FUNCTION_BLOCK FB_LightTower
VAR_INPUT
	bBuzzerBypass: BOOL;
END_VAR
VAR_OUTPUT
	qLedGreen	: BOOL;
	qLedYellow	: BOOL;
	qLedRed		: BOOL;
	qLedBlue	: BOOL;
	qBuzzer		: BOOL;		
	
	qSignal_1: BOOL; //wire BN
	qSignal_2: BOOL; //wire GY
	qSignal_3: BOOL; //wire BK
	qSignal_4: BOOL; //wire WT

END_VAR
VAR
	eLightTowerState		: E_LightTowerState;
	eLightTower_Type		: E_LightTower_Type:=E_LightTower_Type.eSingleLayer;

	
	ton_Blink				: TON;
	ton_Buzzer				: TON;
	t_Buzzer				: TIME:=T#2S;
	t_BuzzerShort			: TIME:=T#0.5S;
	t_BuzzerErrorDelay		: TIME:=T#10S;
	t_BuzzerWarningDelay	: TIME:=T#30S;
	//eLightTowerState_Last	: E_LightTowerState;
	bBuzzerMuteMemo: BOOL;	
	ton_MuteBuzzer: TON;
	ton_NoMessage: TON;
	ton_BuzzerLongTimeOn: TON;	
END_VAR

ton_Blink(IN:=NOT ton_Blink.Q);
CASE eLightTower_Type OF
	E_LightTower_Type.eSingleLayer: m_Single_Layer();
	E_LightTower_Type.eMultiLayer: m_Multi_Layer();
	
END_CASE


ton_NoMessage(PT:=T#5S,IN:=bBuzzerMuteMemo AND iActErrors=0 AND iActWarning=0);

IF (stOpMain.bSetPlay
	(*OR stOpLoad.bSetPlay
	OR stOpUnload.bSetPlay
	OR stOpManip.bSetPlay
	OR stOpHMI.bSetPlay
	OR prg_Call_OpMode.fbModeIndex.rt_Play.Q
	OR prg_Call_OpMode.fbModeLoad.rt_Play.Q
	OR prg_Call_OpMode.fbModeUnload.rt_Play.Q
	OR prg_Call_OpMode.fbModeManip.rt_Play.Q*)
	OR ton_NoMessage.Q	
)
THEN;
	ton_MuteBuzzer.IN:=TRUE;
END_IF
IF ton_MuteBuzzer.IN THEN;
	bBuzzerMuteMemo:=FALSE;
END_IF
ton_MuteBuzzer(PT:=T#1S);
IF ton_MuteBuzzer.Q THEN
	ton_MuteBuzzer.IN:=FALSE;
END_IF
IF prg_Messages.ResetErrors OR ton_BuzzerLongTimeOn.Q THEN;// iActErrors=0 AND iActWarning=0
	bBuzzerMuteMemo:=TRUE;
END_IF
ton_BuzzerLongTimeOn(PT:=T#30M,IN:=eBuzzerMode<>eBuzzerOff);

(*
TYPE E_BuzzerMode :
(
	eBuzzerOff := 0,
	eBuzzerError,		//Short Delay Off
	eBuzzerWarning		//Long Delay Off
);
END_TYPE
*)

IF NOT bBuzzerBypass THEN
	ton_Buzzer();
	CASE eBuzzerMode OF
		eBuzzerOff :;
			qBuzzer:=FALSE;
			
			ton_Buzzer.IN:=FALSE;
		eBuzzerError:;			//Short Delay Off
			qBuzzer:=TRUE;
			ton_Buzzer.PT:=t_BuzzerErrorDelay;
			ton_Buzzer.IN:=NOT ton_Buzzer.Q;
			IF ton_Buzzer.ET>t_Buzzer THEN; qBuzzer:=FALSE; END_IF
		eBuzzerWarning:;		//Long Delay Off
			qBuzzer:=TRUE;
			ton_Buzzer.PT:=t_BuzzerWarningDelay;
			ton_Buzzer.IN:=NOT ton_Buzzer.Q;
			IF ton_Buzzer.ET>t_BuzzerShort THEN; qBuzzer:=FALSE; END_IF
	END_CASE	
ELSE
	qBuzzer:=FALSE;
END_IF

METHOD m_Multi_Layer : BOOL
VAR_INPUT
END_VAR
CASE eLightTowerState OF
	E_LightTowerState.eLightsOff:;
		qLedGreen	:=FALSE;
		qLedYellow	:=FALSE;
		qLedRed		:=FALSE;
		qLedBlue	:=FALSE;
		eBuzzerMode:=eBuzzerOff;	
		
	E_LightTowerState.eGreen:;
		qLedGreen	:=TRUE;
		qLedYellow	:=FALSE;
		qLedRed		:=FALSE;
		qLedBlue	:=FALSE;
		eBuzzerMode:=eBuzzerOff;	
		
	E_LightTowerState.eGreen_YellowBlink:;
		qLedGreen	:=TRUE;
		qLedYellow	:=TRUE;
		qLedRed		:=FALSE;
		qLedBlue	:=FALSE;
		IF bBuzzerMuteMemo THEN;
			eBuzzerMode:=eBuzzerOff;
		ELSE
			eBuzzerMode:=eBuzzerWarning;
		END_IF
		ton_Blink.PT:=T#1S;
		IF ton_Blink.ET>T#0.5S THEN; qLedYellow:=FALSE; ELSE;qLedGreen:=FALSE; END_IF	
		
	E_LightTowerState.eGreenBlink:;
		qLedGreen	:=TRUE;
		qLedYellow	:=FALSE;
		qLedRed		:=FALSE;
		qLedBlue	:=FALSE;
		eBuzzerMode:=eBuzzerOff;		
		ton_Blink.PT:=T#1S;
		IF ton_Blink.ET>T#0.5S THEN; qLedGreen:=FALSE; END_IF	

	E_LightTowerState.eGreenBlink_YellowBlink:;
		qLedGreen	:=TRUE;
		qLedYellow	:=TRUE;
		qLedRed		:=FALSE;
		qLedBlue	:=FALSE;
		IF bBuzzerMuteMemo THEN;
			eBuzzerMode:=eBuzzerOff;
		ELSE
			eBuzzerMode:=eBuzzerWarning;
		END_IF
		ton_Blink.PT:=T#1S;
		IF ton_Blink.ET>T#0.5S THEN; qLedYellow:=FALSE; ELSE;qLedGreen:=FALSE; END_IF

	E_LightTowerState.eGreenBlink_RedBlink:;
		qLedGreen	:=TRUE;
		qLedYellow	:=FALSE;
		qLedRed		:=TRUE;
		qLedBlue	:=FALSE;
		IF bBuzzerMuteMemo THEN;
			eBuzzerMode:=eBuzzerOff;
		ELSE
			eBuzzerMode:=eBuzzerError;
		END_IF
		ton_Blink.PT:=T#1S;
		IF ton_Blink.ET>T#0.5S THEN; qLedRed:=FALSE; ELSE;qLedGreen:=FALSE; END_IF
		
	E_LightTowerState.eYellow:;
		qLedGreen	:=FALSE;
		qLedYellow	:=TRUE;
		qLedRed		:=FALSE;
		qLedBlue	:=FALSE;
		eBuzzerMode:=eBuzzerOff;	
		
	E_LightTowerState.eRed:;
		qLedGreen	:=FALSE;
		qLedYellow	:=FALSE;
		qLedRed		:=TRUE;
		qLedBlue	:=FALSE;
		IF bBuzzerMuteMemo THEN;
			eBuzzerMode:=eBuzzerOff;
		ELSE
			eBuzzerMode:=eBuzzerError;
		END_IF
		
	E_LightTowerState.eBlue:;
		qLedGreen	:=FALSE;
		qLedYellow	:=FALSE;
		qLedRed		:=FALSE;
		qLedBlue	:=TRUE;
		eBuzzerMode:=eBuzzerOff;	
				
END_CASE
END_METHOD

METHOD m_Op_Case1 : BOOL
VAR_INPUT
END_VAR
IF 		stOpMain.iActOperation=E_OperationButtons.ePauseAll
	AND iActErrors<>0
	THEN;	
	eLightTowerState:=E_LightTowerState.eRed;
 						//7
ELSIF 	stOpMain.iActOperation=E_OperationButtons.ePauseAll
	AND iActErrors=0
	THEN;
	eLightTowerState:=E_LightTowerState.eYellow;					//6	
	
ELSIF 	stOpMain.iActOperation=E_OperationButtons.ePlayAll
	AND iActErrors=0
 	AND iActWarning<>0
	THEN;
	eLightTowerState:=E_LightTowerState.eGreenBlink_YellowBlink;	//4
		
ELSIF 	stOpMain.iActOperation=E_OperationButtons.ePlayAll
	AND iActErrors=0 
	AND iActWarning=0 
	THEN;
	eLightTowerState:=E_LightTowerState.eGreen;						//1
END_IF
END_METHOD

METHOD m_Op_Case2 : BOOL
VAR_INPUT
END_VAR
IF 		stOpMain.iActOperation=E_OperationButtons.ePauseAll
	//AND stOpLoad.iActOperation=E_OperationButtons.ePauseAll
	//AND stOpUnload.iActOperation=E_OperationButtons.ePauseAll
	//AND stOpManip.iActOperation=E_OperationButtons.ePauseAll
	//AND stOpHMI.iActOperation=E_OperationButtons.ePauseAll
	AND iActErrors<>0
	THEN;	
	eLightTowerState:=E_LightTowerState.eRed;
 						//7
ELSIF 	stOpMain.iActOperation=E_OperationButtons.ePauseAll
	//AND stOpLoad.iActOperation=E_OperationButtons.ePauseAll
	//AND stOpUnload.iActOperation=E_OperationButtons.ePauseAll
	//AND stOpManip.iActOperation=E_OperationButtons.ePauseAll
	//AND stOpHMI.iActOperation=E_OperationButtons.ePauseAll
	AND iActErrors=0
	THEN;
	eLightTowerState:=E_LightTowerState.eYellow;					//6
	
ELSIF 	(stOpMain.iActOperation=E_OperationButtons.ePlayAll
	(*OR stOpLoad.iActOperation=E_OperationButtons.ePlayAll
	OR stOpUnload.iActOperation=E_OperationButtons.ePlayAll
	OR stOpManip.iActOperation=E_OperationButtons.ePlayAll
	OR stOpHMI.iActOperation=E_OperationButtons.ePlayAll*))
	AND iActErrors<>0 
	THEN;
	eLightTowerState:=E_LightTowerState.eGreenBlink_RedBlink;		//5
	
ELSIF 	(stOpMain.iActOperation=E_OperationButtons.ePlayAll
	(*OR stOpLoad.iActOperation=E_OperationButtons.ePlayAll
	OR stOpUnload.iActOperation=E_OperationButtons.ePlayAll
	OR stOpManip.iActOperation=E_OperationButtons.ePlayAll
	OR stOpHMI.iActOperation=E_OperationButtons.ePlayAll*))
	AND iActErrors=0
 	AND iActWarning<>0
	THEN;
	eLightTowerState:=E_LightTowerState.eGreenBlink_YellowBlink;	//4
	
ELSIF  	(stOpMain.iActOperation=E_OperationButtons.ePlayAll
	(*OR stOpLoad.iActOperation=E_OperationButtons.ePlayAll
	OR stOpUnload.iActOperation=E_OperationButtons.ePlayAll
	OR stOpManip.iActOperation=E_OperationButtons.ePlayAll
	OR stOpHMI.iActOperation=E_OperationButtons.ePlayAll*))
	AND  (stOpMain.iActOperation=E_OperationButtons.ePauseAll
	(*OR stOpLoad.iActOperation=E_OperationButtons.ePauseAll
	OR stOpUnload.iActOperation=E_OperationButtons.ePauseAll
	OR stOpManip.iActOperation=E_OperationButtons.ePauseAll
	OR stOpHMI.iActOperation=E_OperationButtons.ePauseAll*))	
	AND iActErrors=0
 	AND iActWarning=0
	THEN;
	eLightTowerState:=E_LightTowerState.eGreenBlink;				//3
	
ELSIF 	stOpMain.iActOperation=E_OperationButtons.ePlayAll
	(*AND stOpLoad.iActOperation=E_OperationButtons.ePlayAll
	AND stOpUnload.iActOperation=E_OperationButtons.ePlayAll
	AND stOpManip.iActOperation=E_OperationButtons.ePlayAll
	AND stOpHMI.iActOperation=E_OperationButtons.ePlayAll*)
	AND iActErrors=0 
	AND iActWarning<>0
	THEN;
	eLightTowerState:=E_LightTowerState.eGreen_YellowBlink;			//2
	
ELSIF 	stOpMain.iActOperation=E_OperationButtons.ePlayAll
	(*AND stOpLoad.iActOperation=E_OperationButtons.ePlayAll
	AND stOpUnload.iActOperation=E_OperationButtons.ePlayAll
	AND stOpManip.iActOperation=E_OperationButtons.ePlayAll
	AND stOpHMI.iActOperation=E_OperationButtons.ePlayAll*)
	AND iActErrors=0 
	AND iActWarning=0 
	THEN;
	eLightTowerState:=E_LightTowerState.eGreen;						//1
END_IF
END_METHOD

METHOD m_Op_Case3 : BOOL
VAR_INPUT
END_VAR
END_METHOD

METHOD m_Single_Layer : BOOL
VAR_INPUT
END_VAR
CASE eLightTowerState OF
	E_LightTowerState.eLightsOff:;
		qLedGreen	:=FALSE;
		qLedYellow	:=FALSE;
		qLedRed		:=FALSE;
		qLedBlue	:=FALSE;
		eBuzzerMode:=eBuzzerOff;	
		
	E_LightTowerState.eGreen:;
		qLedGreen	:=TRUE;
		qLedYellow	:=FALSE;
		qLedRed		:=FALSE;
		qLedBlue	:=FALSE;
		eBuzzerMode:=eBuzzerOff;	
		
	E_LightTowerState.eGreen_YellowBlink:;
		qLedGreen	:=TRUE;
		qLedYellow	:=TRUE;
		qLedRed		:=FALSE;
		qLedBlue	:=FALSE;
		IF bBuzzerMuteMemo THEN;
			eBuzzerMode:=eBuzzerOff;
		ELSE
			eBuzzerMode:=eBuzzerWarning;
		END_IF
		ton_Blink.PT:=T#1S;
		IF ton_Blink.ET>T#0.5S THEN; qLedYellow:=FALSE; ELSE;qLedGreen:=FALSE; END_IF	
		
	E_LightTowerState.eGreenBlink:;
		qLedGreen	:=TRUE;
		qLedYellow	:=FALSE;
		qLedRed		:=FALSE;
		qLedBlue	:=FALSE;
		eBuzzerMode:=eBuzzerOff;		
		ton_Blink.PT:=T#1S;
		IF ton_Blink.ET>T#0.5S THEN; qLedGreen:=FALSE; END_IF	

	E_LightTowerState.eGreenBlink_YellowBlink:;
		qLedGreen	:=TRUE;
		qLedYellow	:=TRUE;
		qLedRed		:=FALSE;
		qLedBlue	:=FALSE;
		IF bBuzzerMuteMemo THEN;
			eBuzzerMode:=eBuzzerOff;
		ELSE
			eBuzzerMode:=eBuzzerWarning;
		END_IF
		ton_Blink.PT:=T#1S;
		IF ton_Blink.ET>T#0.5S THEN; qLedYellow:=FALSE; ELSE;qLedGreen:=FALSE; END_IF

	E_LightTowerState.eGreenBlink_RedBlink:;
		qLedGreen	:=TRUE;
		qLedYellow	:=FALSE;
		qLedRed		:=TRUE;
		qLedBlue	:=FALSE;
		IF bBuzzerMuteMemo THEN;
			eBuzzerMode:=eBuzzerOff;
		ELSE
			eBuzzerMode:=eBuzzerError;
		END_IF
		ton_Blink.PT:=T#1S;
		IF ton_Blink.ET>T#0.5S THEN; qLedRed:=FALSE; ELSE;qLedGreen:=FALSE; END_IF
		
	E_LightTowerState.eYellow:;
		qLedGreen	:=FALSE;
		qLedYellow	:=TRUE;
		qLedRed		:=FALSE;
		qLedBlue	:=FALSE;
		eBuzzerMode:=eBuzzerOff;	
		
	E_LightTowerState.eRed:;
		qLedGreen	:=FALSE;
		qLedYellow	:=FALSE;
		qLedRed		:=TRUE;
		qLedBlue	:=FALSE;
		IF bBuzzerMuteMemo THEN;
			eBuzzerMode:=eBuzzerOff;
		ELSE
			eBuzzerMode:=eBuzzerError;
		END_IF
		
	E_LightTowerState.eBlue:;
		qLedGreen	:=FALSE;
		qLedYellow	:=FALSE;
		qLedRed		:=FALSE;
		qLedBlue	:=TRUE;
		eBuzzerMode:=eBuzzerOff;	
				
END_CASE


IF qLedRed THEN;
	qSignal_1:=TRUE;	//wire BN
	qSignal_2:=FALSE;	//wire GY
	qSignal_3:=FALSE;	//wire BK
	qSignal_4:=FALSE;	//wire WT	
ELSIF qLedYellow THEN;
	qSignal_1:=TRUE;	//wire BN
	qSignal_2:=FALSE;	//wire GY
	qSignal_3:=FALSE;	//wire BK
	qSignal_4:=TRUE;	//wire WT	
ELSIF qLedGreen THEN;
	qSignal_1:=FALSE;	//wire BN
	qSignal_2:=FALSE;	//wire GY
	qSignal_3:=FALSE;	//wire BK
	qSignal_4:=TRUE;	//wire WT	
ELSIF qLedBlue THEN;
	qSignal_1:=FALSE;	//wire BN
	qSignal_2:=TRUE;	//wire GY
	qSignal_3:=FALSE;	//wire BK
	qSignal_4:=FALSE;	//wire WT	
ELSE;
	qSignal_1:=FALSE;	//wire BN
	qSignal_2:=FALSE;	//wire GY
	qSignal_3:=FALSE;	//wire BK
	qSignal_4:=FALSE;	//wire WT
END_IF
END_METHOD

PROPERTY pState : E_LightTowerState
GET
pState:=eLightTowerState;
END_GET
SET
eLightTowerState:=pState;
END_SET
END_PROPERTY

END_FUNCTION_BLOCK

(* stored: Version 1.1.0.1, ProductVersion 3.1.4024.15
   POU FB_LightTower: Id {d6cadccd-9ab2-46a9-9355-0d0444ba0b75}, SpecialFunc None
   Method m_Multi_Layer: Id {f813da95-f288-460b-9d28-4c9b377be341}
   Method m_Op_Case1: Id {a6b18087-02cb-4fbe-87dc-e00d38ec9f3d}
   Method m_Op_Case2: Id {6beab5aa-13b0-4367-9a27-d87b42c9f182}
   Method m_Op_Case3: Id {535e2ede-5d19-410d-a152-9f18138e3307}
   Method m_Single_Layer: Id {807e5bcf-8516-486e-b821-87be2aad51ac}
   Property pState: Id {88d147a0-4679-47f6-a24a-a7b90f823d80}
   Get Get: Id {40bac962-88f1-4e9f-ac5e-956f192760cd}
   Set Set: Id {6db856c8-700b-4b17-af46-01ec428eba79} *)
